Fanuc KAREL source: kd00036.KL

-- PROVISIONAL review KL for V770-1; original PC SHA256 7e2ab9476625ff02eae78131e51a01ab69c574e5dbfbd67414c0ed24d64e8817
-- Incomplete behavior may be omitted. Consult companion uncertainty JSON. Do not deploy.
PROGRAM KD00036
%NOLOCKGROUP
VAR
  I : INTEGER
  J : INTEGER
  B : BOOLEAN
  R : REAL
  S : STRING[80]
BEGIN
  -- UNRESOLVED_PC offsets 5-17; opcodes 9D,81,18,9D,1B,9D,12,13,04
  -- UNRESOLVED_PC offsets 22-26; opcodes 7F
END KD00036
